Fanuc KAREL source: kt00008.KL

-- PROVISIONAL review KL for V770-1; original PC SHA256 20967a45cddf9140f831c92bec78f584e640c32018afe5d89a0ab258fc172fb2
-- Incomplete behavior may be omitted. Consult companion uncertainty JSON. Do not deploy.
PROGRAM KT00008
%NOLOCKGROUP
VAR
  I1 : INTEGER
  OUT : REAL
-- UNRESOLVED_DECL H2 type=002017
BEGIN
  -- UNRESOLVED_PC offsets 5-16; opcodes 2E,23
  -- UNRESOLVED_PC offsets 21-35; opcodes 2E,22,9D,33,B4
  -- UNRESOLVED_PC offsets 40-63; opcodes 21,22,9D,33,B3,52,64,23
  -- UNRESOLVED_PC offsets 68-72; opcodes 7F
END KT00008
